// TIA Portal V15.1 export
// export: Created 2026-11-01T00:00:00Z, ExportSetting WithDefaults
Screen "Alarms"  480x272, Number=5, Template=Template_1
  ScreenLayer 
    Rectangle "Rectangle_1" at 0,0 size 480x26
    TextField "Text_1" at 6,2 size 300x22  Text="LCP-01 Alarms"
    TextField "Text_2" at 330,3 size 146x20  Text="E-STOP / RESET"
      SingleBitVisibilityAnimation "VisibilityAnimation"
        tag Sys_Alm_EStop
    Button "Button_1" at 2,236 size 76x34  Mode=Text, TextOff="Overview", TextOn="Overview"
      on Press: ActivateScreen(Screen name := Root screen, Object number := 0)
    Button "Button_2" at 82,236 size 76x34  Mode=Text, TextOff="BR01", TextOn="BR01"
      on Press: ActivateScreen(Screen name := BR01, Object number := 0)
    Button "Button_3" at 162,236 size 76x34  Mode=Text, TextOff="BR02", TextOn="BR02"
      on Press: ActivateScreen(Screen name := BR02, Object number := 0)
    Button "Button_4" at 242,236 size 76x34  Mode=Text, TextOff="Scrubber", TextOn="Scrubber"
      on Press: ActivateScreen(Screen name := Scrubber, Object number := 0)
    Button "Button_5" at 322,236 size 76x34  Mode=Text, TextOff="Alarms", TextOn="Alarms"
      on Press: ActivateScreen(Screen name := Alarms, Object number := 0)
    Button "Button_6" at 402,236 size 76x34  Mode=Text, TextOff="Settings", TextOn="Settings"
      on Press: ActivateScreen(Screen name := Settings, Object number := 0)
    Rectangle "Rectangle_2" at 4,30 size 472x202
    TextField "Text_3" at 12,110 size 456x40  Text="Alarm view goes here (placed by hand in TIA, 0007 P6)"
